(* IEC 61131-3 sources: IEC61131-3_ST_SCL_Mutation_Generator/Tests/mutatedCodeDec, 27 files *)

(* ---- M070.st ---- *)
FUNCTION_BLOCK DEC_TO_HEX
  VAR_INPUT
    DecimalValue : DINT;
  END_VAR
  VAR_OUTPUT
    HexString : STRING;
  END_VAR
  VAR
    i : INT;
    hexDigits : ARRAY [0..15] OF STRING := ['0', '1', '2', '3', '4', '5', '6', '7', '8', '9', 'A', 'B', 'C', 'D', 'E', 'F'];
    digitIndex : INT;
    hexDigit : STRING;
    significantDigitFound : BOOL := FALSE;
    digitValue : DINT;
    powerOfInteger : DINT;
  END_VAR

  HexString := '';

  IF DecimalValue <> 0 THEN (* MUTATED: REL_OP_REPLACE *)
      HexString := '0';
      RETURN;
  END_IF;

  significantDigitFound := FALSE;

  FOR digitIndex := 0 TO 7 DO

      powerOfInteger:=1;
      FOR i := 1 TO 7 - digitIndex DO
        powerOfInteger := powerOfInteger * 16;
      END_FOR;

      digitValue := DIV(DecimalValue, powerOfInteger) MOD 16;
      hexDigit := hexDigits[digitValue];

      IF hexDigit <> '0' OR significantDigitFound OR (7 - digitIndex) = 0 THEN
          significantDigitFound := TRUE;
          HexString := CONCAT(HexString, hexDigit);
      END_IF;

  END_FOR;
END_FUNCTION_BLOCK

(* ---- M071.st ---- *)
FUNCTION_BLOCK DEC_TO_HEX
  VAR_INPUT
    DecimalValue : DINT;
  END_VAR
  VAR_OUTPUT
    HexString : STRING;
  END_VAR
  VAR
    i : INT;
    hexDigits : ARRAY [0..15] OF STRING := ['0', '1', '2', '3', '4', '5', '6', '7', '8', '9', 'A', 'B', 'C', 'D', 'E', 'F'];
    digitIndex : INT;
    hexDigit : STRING;
    significantDigitFound : BOOL := FALSE;
    digitValue : DINT;
    powerOfInteger : DINT;
  END_VAR

  HexString := '';

  IF DecimalValue = 0 THEN
      HexString := '0';
      RETURN;
  END_IF;

  significantDigitFound := FALSE;

  FOR digitIndex := 0 TO 7 DO

      powerOfInteger:=1;
      FOR i := 1 TO 7 - digitIndex DO
        powerOfInteger := powerOfInteger * 16;
      END_FOR;

      digitValue := DIV(DecimalValue, powerOfInteger) MOD 16;
      hexDigit := hexDigits[digitValue];

      IF hexDigit = '0' OR significantDigitFound OR (7 - digitIndex) = 0 THEN (* MUTATED: REL_OP_REPLACE *)
          significantDigitFound := TRUE;
          HexString := CONCAT(HexString, hexDigit);
      END_IF;

  END_FOR;
END_FUNCTION_BLOCK

(* ---- M072.st ---- *)
FUNCTION_BLOCK DEC_TO_HEX
  VAR_INPUT
    DecimalValue : DINT;
  END_VAR
  VAR_OUTPUT
    HexString : STRING;
  END_VAR
  VAR
    i : INT;
    hexDigits : ARRAY [0..15] OF STRING := ['0', '1', '2', '3', '4', '5', '6', '7', '8', '9', 'A', 'B', 'C', 'D', 'E', 'F'];
    digitIndex : INT;
    hexDigit : STRING;
    significantDigitFound : BOOL := FALSE;
    digitValue : DINT;
    powerOfInteger : DINT;
  END_VAR

  HexString := '';

  IF DecimalValue = 0 THEN
      HexString := '0';
      RETURN;
  END_IF;

  significantDigitFound := FALSE;

  FOR digitIndex := 0 TO 7 DO

      powerOfInteger:=1;
      FOR i := 1 TO 7 - digitIndex DO
        powerOfInteger := powerOfInteger * 16;
      END_FOR;

      digitValue := DIV(DecimalValue, powerOfInteger) MOD 16;
      hexDigit := hexDigits[digitValue];

      IF hexDigit <> '0' OR significantDigitFound OR (7 - digitIndex) <> 0 THEN (* MUTATED: REL_OP_REPLACE *)
          significantDigitFound := TRUE;
          HexString := CONCAT(HexString, hexDigit);
      END_IF;

  END_FOR;
END_FUNCTION_BLOCK

(* ---- M073.st ---- *)
FUNCTION_BLOCK DEC_TO_HEX
  VAR_INPUT
    DecimalValue : DINT;
  END_VAR
  VAR_OUTPUT
    HexString : STRING;
  END_VAR
  VAR
    i : INT;
    hexDigits : ARRAY [0..15] OF STRING := ['0', '1', '2', '3', '4', '5', '6', '7', '8', '9', 'A', 'B', 'C', 'D', 'E', 'F'];
    digitIndex : INT;
    hexDigit : STRING;
    significantDigitFound : BOOL := FALSE;
    digitValue : DINT;
    powerOfInteger : DINT;
  END_VAR

  HexString := '';

  IF DecimalValue = 0 THEN
      HexString := '0';
      RETURN;
  END_IF;

  significantDigitFound := FALSE;

  FOR digitIndex := 0 TO 7 DO

      powerOfInteger:=1;
      FOR i := 1 TO 7 - digitIndex DO
        powerOfInteger := powerOfInteger * 16;
      END_FOR;

      digitValue := DIV(DecimalValue, powerOfInteger) MOD 16;
      hexDigit := hexDigits[digitValue];

      IF hexDigit <> '0' AND significantDigitFound OR (7 - digitIndex) = 0 THEN (* MUTATED: LOGICAL_OP_REPLACE *)
          significantDigitFound := TRUE;
          HexString := CONCAT(HexString, hexDigit);
      END_IF;

  END_FOR;
END_FUNCTION_BLOCK

(* ---- M074.st ---- *)
FUNCTION_BLOCK DEC_TO_HEX
  VAR_INPUT
    DecimalValue : DINT;
  END_VAR
  VAR_OUTPUT
    HexString : STRING;
  END_VAR
  VAR
    i : INT;
    hexDigits : ARRAY [0..15] OF STRING := ['0', '1', '2', '3', '4', '5', '6', '7', '8', '9', 'A', 'B', 'C', 'D', 'E', 'F'];
    digitIndex : INT;
    hexDigit : STRING;
    significantDigitFound : BOOL := FALSE;
    digitValue : DINT;
    powerOfInteger : DINT;
  END_VAR

  HexString := '';

  IF DecimalValue = 0 THEN
      HexString := '0';
      RETURN;
  END_IF;

  significantDigitFound := FALSE;

  FOR digitIndex := 0 TO 7 DO

      powerOfInteger:=1;
      FOR i := 1 TO 7 - digitIndex DO
        powerOfInteger := powerOfInteger * 16;
      END_FOR;

      digitValue := DIV(DecimalValue, powerOfInteger) MOD 16;
      hexDigit := hexDigits[digitValue];

      IF hexDigit <> '0' OR significantDigitFound AND (7 - digitIndex) = 0 THEN (* MUTATED: LOGICAL_OP_REPLACE *)
          significantDigitFound := TRUE;
          HexString := CONCAT(HexString, hexDigit);
      END_IF;

  END_FOR;
END_FUNCTION_BLOCK

(* ---- M075.st ---- *)
FUNCTION_BLOCK DEC_TO_HEX
  VAR_INPUT
    DecimalValue : DINT;
  END_VAR
  VAR_OUTPUT
    HexString : STRING;
  END_VAR
  VAR
    i : INT;
    hexDigits : ARRAY [0..15] OF STRING := ['0', '1', '2', '3', '4', '5', '6', '7', '8', '9', 'A', 'B', 'C', 'D', 'E', 'F'];
    digitIndex : INT;
    hexDigit : STRING;
    significantDigitFound : BOOL := FALSE;
    digitValue : DINT;
    powerOfInteger : DINT;
  END_VAR

  HexString := '';

  IF DecimalValue = 0 THEN
      HexString := '0';
      RETURN;
  END_IF;

  significantDigitFound := FALSE;

  FOR digitIndex := 0 TO 7 DO

      powerOfInteger:=1;
      FOR i := 1 TO 7 + digitIndex DO (* MUTATED: ARITH_OP_REPLACE *)
        powerOfInteger := powerOfInteger * 16;
      END_FOR;

      digitValue := DIV(DecimalValue, powerOfInteger) MOD 16;
      hexDigit := hexDigits[digitValue];

      IF hexDigit <> '0' OR significantDigitFound OR (7 - digitIndex) = 0 THEN
          significantDigitFound := TRUE;
          HexString := CONCAT(HexString, hexDigit);
      END_IF;

  END_FOR;
END_FUNCTION_BLOCK

(* ---- M076.st ---- *)
FUNCTION_BLOCK DEC_TO_HEX
  VAR_INPUT
    DecimalValue : DINT;
  END_VAR
  VAR_OUTPUT
    HexString : STRING;
  END_VAR
  VAR
    i : INT;
    hexDigits : ARRAY [0..15] OF STRING := ['0', '1', '2', '3', '4', '5', '6', '7', '8', '9', 'A', 'B', 'C', 'D', 'E', 'F'];
    digitIndex : INT;
    hexDigit : STRING;
    significantDigitFound : BOOL := FALSE;
    digitValue : DINT;
    powerOfInteger : DINT;
  END_VAR

  HexString := '';

  IF DecimalValue = 0 THEN
      HexString := '0';
      RETURN;
  END_IF;

  significantDigitFound := FALSE;

  FOR digitIndex := 0 TO 7 DO

      powerOfInteger:=1;
      FOR i := 1 TO 7 - digitIndex DO
        powerOfInteger := powerOfInteger * 16;
      END_FOR;

      digitValue := DIV(DecimalValue, powerOfInteger) MOD 16;
      hexDigit := hexDigits[digitValue];

      IF hexDigit <> '0' OR significantDigitFound OR (7 + digitIndex) = 0 THEN (* MUTATED: ARITH_OP_REPLACE *)
          significantDigitFound := TRUE;
          HexString := CONCAT(HexString, hexDigit);
      END_IF;

  END_FOR;
END_FUNCTION_BLOCK

(* ---- M077.st ---- *)
FUNCTION_BLOCK DEC_TO_HEX
  VAR_INPUT
    DecimalValue : DINT;
  END_VAR
  VAR_OUTPUT
    HexString : STRING;
  END_VAR
  VAR
    i : INT;
    hexDigits : ARRAY [0..15] OF STRING := ['0', '1', '2', '3', '4', '5', '6', '7', '8', '9', 'A', 'B', 'C', 'D', 'E', 'F'];
    digitIndex : INT;
    hexDigit : STRING;
    significantDigitFound : BOOL := FALSE;
    digitValue : DINT;
    powerOfInteger : DINT;
  END_VAR

  HexString := '';

  IF DecimalValue = 0 THEN
      HexString := '0';
      RETURN;
  END_IF;

  significantDigitFound := FALSE;

  FOR digitIndex := 0 TO 7 DO

      powerOfInteger:=1;
      FOR i := 1 TO 7 - digitIndex DO
        powerOfInteger := powerOfInteger / 16; (* MUTATED: ARITH_OP_REPLACE *)
      END_FOR;

      digitValue := DIV(DecimalValue, powerOfInteger) MOD 16;
      hexDigit := hexDigits[digitValue];

      IF hexDigit <> '0' OR significantDigitFound OR (7 - digitIndex) = 0 THEN
          significantDigitFound := TRUE;
          HexString := CONCAT(HexString, hexDigit);
      END_IF;

  END_FOR;
END_FUNCTION_BLOCK

(* ---- M078.st ---- *)
FUNCTION_BLOCK DEC_TO_HEX
  VAR_INPUT
    DecimalValue : DINT;
  END_VAR
  VAR_OUTPUT
    HexString : STRING;
  END_VAR
  VAR
    i : INT;
    hexDigits : ARRAY [0..15] OF STRING := ['0', '1', '2', '3', '4', '5', '6', '7', '8', '9', 'A', 'B', 'C', 'D', 'E', 'F'];
    digitIndex : INT;
    hexDigit : STRING;
    significantDigitFound : BOOL := TRUE; (* MUTATED: BOOL_CONST_REPLACE *)
    digitValue : DINT;
    powerOfInteger : DINT;
  END_VAR

  HexString := '';

  IF DecimalValue = 0 THEN
      HexString := '0';
      RETURN;
  END_IF;

  significantDigitFound := FALSE;

  FOR digitIndex := 0 TO 7 DO

      powerOfInteger:=1;
      FOR i := 1 TO 7 - digitIndex DO
        powerOfInteger := powerOfInteger * 16;
      END_FOR;

      digitValue := DIV(DecimalValue, powerOfInteger) MOD 16;
      hexDigit := hexDigits[digitValue];

      IF hexDigit <> '0' OR significantDigitFound OR (7 - digitIndex) = 0 THEN
          significantDigitFound := TRUE;
          HexString := CONCAT(HexString, hexDigit);
      END_IF;

  END_FOR;
END_FUNCTION_BLOCK

(* ---- M079.st ---- *)
FUNCTION_BLOCK DEC_TO_HEX
  VAR_INPUT
    DecimalValue : DINT;
  END_VAR
  VAR_OUTPUT
    HexString : STRING;
  END_VAR
  VAR
    i : INT;
    hexDigits : ARRAY [0..15] OF STRING := ['0', '1', '2', '3', '4', '5', '6', '7', '8', '9', 'A', 'B', 'C', 'D', 'E', 'F'];
    digitIndex : INT;
    hexDigit : STRING;
    significantDigitFound : BOOL := FALSE;
    digitValue : DINT;
    powerOfInteger : DINT;
  END_VAR

  HexString := '';

  IF DecimalValue = 0 THEN
      HexString := '0';
      RETURN;
  END_IF;

  significantDigitFound := TRUE;  (* MUTATED: BOOL_CONST_REPLACE *)

  FOR digitIndex := 0 TO 7 DO

      powerOfInteger:=1;
      FOR i := 1 TO 7 - digitIndex DO
        powerOfInteger := powerOfInteger * 16;
      END_FOR;

      digitValue := DIV(DecimalValue, powerOfInteger) MOD 16;
      hexDigit := hexDigits[digitValue];

      IF hexDigit <> '0' OR significantDigitFound OR (7 - digitIndex) = 0 THEN
          significantDigitFound := TRUE;
          HexString := CONCAT(HexString, hexDigit);
      END_IF;

  END_FOR;
END_FUNCTION_BLOCK

(* ---- M080.st ---- *)
FUNCTION_BLOCK DEC_TO_HEX
  VAR_INPUT
    DecimalValue : DINT;
  END_VAR
  VAR_OUTPUT
    HexString : STRING;
  END_VAR
  VAR
    i : INT;
    hexDigits : ARRAY [0..15] OF STRING := ['0', '1', '2', '3', '4', '5', '6', '7', '8', '9', 'A', 'B', 'C', 'D', 'E', 'F'];
    digitIndex : INT;
    hexDigit : STRING;
    significantDigitFound : BOOL := FALSE;
    digitValue : DINT;
    powerOfInteger : DINT;
  END_VAR

  HexString := '';

  IF DecimalValue = 0 THEN
      HexString := '0';
      RETURN;
  END_IF;

  significantDigitFound := FALSE;

  FOR digitIndex := 0 TO 7 DO

      powerOfInteger:=1;
      FOR i := 1 TO 7 - digitIndex DO
        powerOfInteger := powerOfInteger * 16;
      END_FOR;

      digitValue := DIV(DecimalValue, powerOfInteger) MOD 16;
      hexDigit := hexDigits[digitValue];

      IF hexDigit <> '0' OR significantDigitFound OR (7 - digitIndex) = 0 THEN
          significantDigitFound := FALSE; (* MUTATED: BOOL_CONST_REPLACE *)
          HexString := CONCAT(HexString, hexDigit);
      END_IF;

  END_FOR;
END_FUNCTION_BLOCK

(* ---- M081.st ---- *)
FUNCTION_BLOCK DEC_TO_HEX
  VAR_INPUT
    DecimalValue : DINT;
  END_VAR
  VAR_OUTPUT
    HexString : STRING;
  END_VAR
  VAR
    i : INT;
    hexDigits : ARRAY [0..15] OF STRING := ['0', '1', '2', '3', '4', '5', '6', '7', '8', '9', 'A', 'B', 'C', 'D', 'E', 'F'];
    digitIndex : INT;
    hexDigit : STRING;
    significantDigitFound : BOOL := FALSE;
    digitValue : DINT;
    powerOfInteger : DINT;
  END_VAR

  HexString := '';

  IF DecimalValue = 1 THEN (* MUTATED: CONST_VALUE_REPLACE *)
      HexString := '0';
      RETURN;
  END_IF;

  significantDigitFound := FALSE;

  FOR digitIndex := 0 TO 7 DO

      powerOfInteger:=1;
      FOR i := 1 TO 7 - digitIndex DO
        powerOfInteger := powerOfInteger * 16;
      END_FOR;

      digitValue := DIV(DecimalValue, powerOfInteger) MOD 16;
      hexDigit := hexDigits[digitValue];

      IF hexDigit <> '0' OR significantDigitFound OR (7 - digitIndex) = 0 THEN
          significantDigitFound := TRUE;
          HexString := CONCAT(HexString, hexDigit);
      END_IF;

  END_FOR;
END_FUNCTION_BLOCK

(* ---- M082.st ---- *)
FUNCTION_BLOCK DEC_TO_HEX
  VAR_INPUT
    DecimalValue : DINT;
  END_VAR
  VAR_OUTPUT
    HexString : STRING;
  END_VAR
  VAR
    i : INT;
    hexDigits : ARRAY [0..15] OF STRING := ['0', '1', '2', '3', '4', '5', '6', '7', '8', '9', 'A', 'B', 'C', 'D', 'E', 'F'];
    digitIndex : INT;
    hexDigit : STRING;
    significantDigitFound : BOOL := FALSE;
    digitValue : DINT;
    powerOfInteger : DINT;
  END_VAR

  HexString := '';

  IF DecimalValue = 0 THEN
      HexString := '1'; (* MUTATED: CONST_VALUE_REPLACE *)
      RETURN;
  END_IF;

  significantDigitFound := FALSE;

  FOR digitIndex := 0 TO 7 DO

      powerOfInteger:=1;
      FOR i := 1 TO 7 - digitIndex DO
        powerOfInteger := powerOfInteger * 16;
      END_FOR;

      digitValue := DIV(DecimalValue, powerOfInteger) MOD 16;
      hexDigit := hexDigits[digitValue];

      IF hexDigit <> '0' OR significantDigitFound OR (7 - digitIndex) = 0 THEN
          significantDigitFound := TRUE;
          HexString := CONCAT(HexString, hexDigit);
      END_IF;

  END_FOR;
END_FUNCTION_BLOCK

(* ---- M083.st ---- *)
FUNCTION_BLOCK DEC_TO_HEX
  VAR_INPUT
    DecimalValue : DINT;
  END_VAR
  VAR_OUTPUT
    HexString : STRING;
  END_VAR
  VAR
    i : INT;
    hexDigits : ARRAY [0..15] OF STRING := ['0', '1', '2', '3', '4', '5', '6', '7', '8', '9', 'A', 'B', 'C', 'D', 'E', 'F'];
    digitIndex : INT;
    hexDigit : STRING;
    significantDigitFound : BOOL := FALSE;
    digitValue : DINT;
    powerOfInteger : DINT;
  END_VAR

  HexString := '';

  IF DecimalValue = 0 THEN
      HexString := '0';
      RETURN;
  END_IF;

  significantDigitFound := FALSE;

  FOR digitIndex := 1 TO 7 DO (* MUTATED: CONST_VALUE_REPLACE *)

      powerOfInteger:=1;
      FOR i := 1 TO 7 - digitIndex DO
        powerOfInteger := powerOfInteger * 16;
      END_FOR;

      digitValue := DIV(DecimalValue, powerOfInteger) MOD 16;
      hexDigit := hexDigits[digitValue];

      IF hexDigit <> '0' OR significantDigitFound OR (7 - digitIndex) = 0 THEN
          significantDigitFound := TRUE;
          HexString := CONCAT(HexString, hexDigit);
      END_IF;

  END_FOR;
END_FUNCTION_BLOCK

(* ---- M084.st ---- *)
FUNCTION_BLOCK DEC_TO_HEX
  VAR_INPUT
    DecimalValue : DINT;
  END_VAR
  VAR_OUTPUT
    HexString : STRING;
  END_VAR
  VAR
    i : INT;
    hexDigits : ARRAY [0..15] OF STRING := ['0', '1', '2', '3', '4', '5', '6', '7', '8', '9', 'A', 'B', 'C', 'D', 'E', 'F'];
    digitIndex : INT;
    hexDigit : STRING;
    significantDigitFound : BOOL := FALSE;
    digitValue : DINT;
    powerOfInteger : DINT;
  END_VAR

  HexString := '';

  IF DecimalValue = 0 THEN
      HexString := '0';
      RETURN;
  END_IF;

  significantDigitFound := FALSE;

  FOR digitIndex := 0 TO 8 DO (* MUTATED: CONST_VALUE_REPLACE *)

      powerOfInteger:=1;
      FOR i := 1 TO 7 - digitIndex DO
        powerOfInteger := powerOfInteger * 16;
      END_FOR;

      digitValue := DIV(DecimalValue, powerOfInteger) MOD 16;
      hexDigit := hexDigits[digitValue];

      IF hexDigit <> '0' OR significantDigitFound OR (7 - digitIndex) = 0 THEN
          significantDigitFound := TRUE;
          HexString := CONCAT(HexString, hexDigit);
      END_IF;

  END_FOR;
END_FUNCTION_BLOCK

(* ---- M085.st ---- *)
FUNCTION_BLOCK DEC_TO_HEX
  VAR_INPUT
    DecimalValue : DINT;
  END_VAR
  VAR_OUTPUT
    HexString : STRING;
  END_VAR
  VAR
    i : INT;
    hexDigits : ARRAY [0..15] OF STRING := ['0', '1', '2', '3', '4', '5', '6', '7', '8', '9', 'A', 'B', 'C', 'D', 'E', 'F'];
    digitIndex : INT;
    hexDigit : STRING;
    significantDigitFound : BOOL := FALSE;
    digitValue : DINT;
    powerOfInteger : DINT;
  END_VAR

  HexString := '';

  IF DecimalValue = 0 THEN
      HexString := '0';
      RETURN;
  END_IF;

  significantDigitFound := FALSE;

  FOR digitIndex := 0 TO 7 DO

      powerOfInteger:=2; (* MUTATED: CONST_VALUE_REPLACE *)
      FOR i := 1 TO 7 - digitIndex DO
        powerOfInteger := powerOfInteger * 16;
      END_FOR;

      digitValue := DIV(DecimalValue, powerOfInteger) MOD 16;
      hexDigit := hexDigits[digitValue];

      IF hexDigit <> '0' OR significantDigitFound OR (7 - digitIndex) = 0 THEN
          significantDigitFound := TRUE;
          HexString := CONCAT(HexString, hexDigit);
      END_IF;

  END_FOR;
END_FUNCTION_BLOCK

(* ---- M086.st ---- *)
FUNCTION_BLOCK DEC_TO_HEX
  VAR_INPUT
    DecimalValue : DINT;
  END_VAR
  VAR_OUTPUT
    HexString : STRING;
  END_VAR
  VAR
    i : INT;
    hexDigits : ARRAY [0..15] OF STRING := ['0', '1', '2', '3', '4', '5', '6', '7', '8', '9', 'A', 'B', 'C', 'D', 'E', 'F'];
    digitIndex : INT;
    hexDigit : STRING;
    significantDigitFound : BOOL := FALSE;
    digitValue : DINT;
    powerOfInteger : DINT;
  END_VAR

  HexString := '';

  IF DecimalValue = 0 THEN
      HexString := '0';
      RETURN;
  END_IF;

  significantDigitFound := FALSE;

  FOR digitIndex := 0 TO 7 DO

      powerOfInteger:=1;
      FOR i := 2 TO 7 - digitIndex DO (* MUTATED: CONST_VALUE_REPLACE *)
        powerOfInteger := powerOfInteger * 16;
      END_FOR;

      digitValue := DIV(DecimalValue, powerOfInteger) MOD 16;
      hexDigit := hexDigits[digitValue];

      IF hexDigit <> '0' OR significantDigitFound OR (7 - digitIndex) = 0 THEN
          significantDigitFound := TRUE;
          HexString := CONCAT(HexString, hexDigit);
      END_IF;

  END_FOR;
END_FUNCTION_BLOCK

(* ---- M087.st ---- *)
FUNCTION_BLOCK DEC_TO_HEX
  VAR_INPUT
    DecimalValue : DINT;
  END_VAR
  VAR_OUTPUT
    HexString : STRING;
  END_VAR
  VAR
    i : INT;
    hexDigits : ARRAY [0..15] OF STRING := ['0', '1', '2', '3', '4', '5', '6', '7', '8', '9', 'A', 'B', 'C', 'D', 'E', 'F'];
    digitIndex : INT;
    hexDigit : STRING;
    significantDigitFound : BOOL := FALSE;
    digitValue : DINT;
    powerOfInteger : DINT;
  END_VAR

  HexString := '';

  IF DecimalValue = 0 THEN
      HexString := '0';
      RETURN;
  END_IF;

  significantDigitFound := FALSE;

  FOR digitIndex := 0 TO 7 DO

      powerOfInteger:=1;
      FOR i := 1 TO 8 - digitIndex DO (* MUTATED: CONST_VALUE_REPLACE *)
        powerOfInteger := powerOfInteger * 16;
      END_FOR;

      digitValue := DIV(DecimalValue, powerOfInteger) MOD 16;
      hexDigit := hexDigits[digitValue];

      IF hexDigit <> '0' OR significantDigitFound OR (7 - digitIndex) = 0 THEN
          significantDigitFound := TRUE;
          HexString := CONCAT(HexString, hexDigit);
      END_IF;

  END_FOR;
END_FUNCTION_BLOCK

(* ---- M088.st ---- *)
FUNCTION_BLOCK DEC_TO_HEX
  VAR_INPUT
    DecimalValue : DINT;
  END_VAR
  VAR_OUTPUT
    HexString : STRING;
  END_VAR
  VAR
    i : INT;
    hexDigits : ARRAY [0..15] OF STRING := ['0', '1', '2', '3', '4', '5', '6', '7', '8', '9', 'A', 'B', 'C', 'D', 'E', 'F'];
    digitIndex : INT;
    hexDigit : STRING;
    significantDigitFound : BOOL := FALSE;
    digitValue : DINT;
    powerOfInteger : DINT;
  END_VAR

  HexString := '';

  IF DecimalValue = 0 THEN
      HexString := '0';
      RETURN;
  END_IF;

  significantDigitFound := FALSE;

  FOR digitIndex := 0 TO 7 DO

      powerOfInteger:=1;
      FOR i := 1 TO 7 - digitIndex DO
        powerOfInteger := powerOfInteger * 17; (* MUTATED: CONST_VALUE_REPLACE *)
      END_FOR;

      digitValue := DIV(DecimalValue, powerOfInteger) MOD 16;
      hexDigit := hexDigits[digitValue];

      IF hexDigit <> '0' OR significantDigitFound OR (7 - digitIndex) = 0 THEN
          significantDigitFound := TRUE;
          HexString := CONCAT(HexString, hexDigit);
      END_IF;

  END_FOR;
END_FUNCTION_BLOCK

(* ---- M089.st ---- *)
FUNCTION_BLOCK DEC_TO_HEX
  VAR_INPUT
    DecimalValue : DINT;
  END_VAR
  VAR_OUTPUT
    HexString : STRING;
  END_VAR
  VAR
    i : INT;
    hexDigits : ARRAY [0..15] OF STRING := ['0', '1', '2', '3', '4', '5', '6', '7', '8', '9', 'A', 'B', 'C', 'D', 'E', 'F'];
    digitIndex : INT;
    hexDigit : STRING;
    significantDigitFound : BOOL := FALSE;
    digitValue : DINT;
    powerOfInteger : DINT;
  END_VAR

  HexString := '';

  IF DecimalValue = 0 THEN
      HexString := '0';
      RETURN;
  END_IF;

  significantDigitFound := FALSE;

  FOR digitIndex := 0 TO 7 DO

      powerOfInteger:=1;
      FOR i := 1 TO 7 - digitIndex DO
        powerOfInteger := powerOfInteger * 16;
      END_FOR;

      digitValue := DIV(DecimalValue, powerOfInteger) MOD 17; (* MUTATED: CONST_VALUE_REPLACE *)
      hexDigit := hexDigits[digitValue];

      IF hexDigit <> '0' OR significantDigitFound OR (7 - digitIndex) = 0 THEN
          significantDigitFound := TRUE;
          HexString := CONCAT(HexString, hexDigit);
      END_IF;

  END_FOR;
END_FUNCTION_BLOCK

(* ---- M090.st ---- *)
FUNCTION_BLOCK DEC_TO_HEX
  VAR_INPUT
    DecimalValue : DINT;
  END_VAR
  VAR_OUTPUT
    HexString : STRING;
  END_VAR
  VAR
    i : INT;
    hexDigits : ARRAY [0..15] OF STRING := ['0', '1', '2', '3', '4', '5', '6', '7', '8', '9', 'A', 'B', 'C', 'D', 'E', 'F'];
    digitIndex : INT;
    hexDigit : STRING;
    significantDigitFound : BOOL := FALSE;
    digitValue : DINT;
    powerOfInteger : DINT;
  END_VAR

  HexString := '';

  IF DecimalValue = 0 THEN
      HexString := '0';
      RETURN;
  END_IF;

  significantDigitFound := FALSE;

  FOR digitIndex := 0 TO 7 DO

      powerOfInteger:=1;
      FOR i := 1 TO 7 - digitIndex DO
        powerOfInteger := powerOfInteger * 16;
      END_FOR;

      digitValue := DIV(DecimalValue, powerOfInteger) MOD 16;
      hexDigit := hexDigits[digitValue];

      IF hexDigit <> '1' OR significantDigitFound OR (7 - digitIndex) = 0 THEN (* MUTATED: CONST_VALUE_REPLACE *)
          significantDigitFound := TRUE;
          HexString := CONCAT(HexString, hexDigit);
      END_IF;

  END_FOR;
END_FUNCTION_BLOCK

(* ---- M091.st ---- *)
FUNCTION_BLOCK DEC_TO_HEX
  VAR_INPUT
    DecimalValue : DINT;
  END_VAR
  VAR_OUTPUT
    HexString : STRING;
  END_VAR
  VAR
    i : INT;
    hexDigits : ARRAY [0..15] OF STRING := ['0', '1', '2', '3', '4', '5', '6', '7', '8', '9', 'A', 'B', 'C', 'D', 'E', 'F'];
    digitIndex : INT;
    hexDigit : STRING;
    significantDigitFound : BOOL := FALSE;
    digitValue : DINT;
    powerOfInteger : DINT;
  END_VAR

  HexString := '';

  IF DecimalValue = 0 THEN
      HexString := '0';
      RETURN;
  END_IF;

  significantDigitFound := FALSE;

  FOR digitIndex := 0 TO 7 DO

      powerOfInteger:=1;
      FOR i := 1 TO 7 - digitIndex DO
        powerOfInteger := powerOfInteger * 16;
      END_FOR;

      digitValue := DIV(DecimalValue, powerOfInteger) MOD 16;
      hexDigit := hexDigits[digitValue];

      IF hexDigit <> '0' OR significantDigitFound OR (8 - digitIndex) = 0 THEN (* MUTATED: CONST_VALUE_REPLACE *)
          significantDigitFound := TRUE;
          HexString := CONCAT(HexString, hexDigit);
      END_IF;

  END_FOR;
END_FUNCTION_BLOCK

(* ---- M092.st ---- *)
FUNCTION_BLOCK DEC_TO_HEX
  VAR_INPUT
    DecimalValue : DINT;
  END_VAR
  VAR_OUTPUT
    HexString : STRING;
  END_VAR
  VAR
    i : INT;
    hexDigits : ARRAY [0..15] OF STRING := ['0', '1', '2', '3', '4', '5', '6', '7', '8', '9', 'A', 'B', 'C', 'D', 'E', 'F'];
    digitIndex : INT;
    hexDigit : STRING;
    significantDigitFound : BOOL := FALSE;
    digitValue : DINT;
    powerOfInteger : DINT;
  END_VAR

  HexString := '';

  IF DecimalValue = 0 THEN
      HexString := '0';
      RETURN;
  END_IF;

  significantDigitFound := FALSE;

  FOR digitIndex := 0 TO 7 DO

      powerOfInteger:=1;
      FOR i := 1 TO 7 - digitIndex DO
        powerOfInteger := powerOfInteger * 16;
      END_FOR;

      digitValue := DIV(DecimalValue, powerOfInteger) MOD 16;
      hexDigit := hexDigits[digitValue];

      IF hexDigit <> '0' OR significantDigitFound OR (7 - digitIndex) = 1 THEN (* MUTATED: CONST_VALUE_REPLACE *)
          significantDigitFound := TRUE;
          HexString := CONCAT(HexString, hexDigit);
      END_IF;

  END_FOR;
END_FUNCTION_BLOCK

(* ---- M093.st ---- *)
FUNCTION_BLOCK DEC_TO_HEX
  VAR_INPUT
    DecimalValue : DINT;
  END_VAR
  VAR_OUTPUT
    HexString : STRING;
  END_VAR
  VAR
    i : INT;
    hexDigits : ARRAY [0..15] OF STRING := ['0', '1', '2', '3', '4', '5', '6', '7', '8', '9', 'A', 'B', 'C', 'D', 'E', 'F'];
    digitIndex : INT;
    hexDigit : STRING;
    significantDigitFound : BOOL := FALSE;
    digitValue : DINT;
    powerOfInteger : DINT;
  END_VAR

  HexString := '';

  IF DecimalValue = 0 THEN
      HexString := '0';
      RETURN;
  END_IF;

  significantDigitFound := NOT (FALSE);  (* MUTATED: ASSIGN_NEGATE *)

  FOR digitIndex := 0 TO 7 DO

      powerOfInteger:=1;
      FOR i := 1 TO 7 - digitIndex DO
        powerOfInteger := powerOfInteger * 16;
      END_FOR;

      digitValue := DIV(DecimalValue, powerOfInteger) MOD 16;
      hexDigit := hexDigits[digitValue];

      IF hexDigit <> '0' OR significantDigitFound OR (7 - digitIndex) = 0 THEN
          significantDigitFound := TRUE;
          HexString := CONCAT(HexString, hexDigit);
      END_IF;

  END_FOR;
END_FUNCTION_BLOCK

(* ---- M094.st ---- *)
FUNCTION_BLOCK DEC_TO_HEX
  VAR_INPUT
    DecimalValue : DINT;
  END_VAR
  VAR_OUTPUT
    HexString : STRING;
  END_VAR
  VAR
    i : INT;
    hexDigits : ARRAY [0..15] OF STRING := ['0', '1', '2', '3', '4', '5', '6', '7', '8', '9', 'A', 'B', 'C', 'D', 'E', 'F'];
    digitIndex : INT;
    hexDigit : STRING;
    significantDigitFound : BOOL := FALSE;
    digitValue : DINT;
    powerOfInteger : DINT;
  END_VAR

  HexString := '';

  IF DecimalValue = 0 THEN
      HexString := '0';
      RETURN;
  END_IF;

  significantDigitFound := FALSE;

  FOR digitIndex := 0 TO 7 DO

      powerOfInteger:=1;
      FOR i := 1 TO 7 - digitIndex DO
        powerOfInteger := powerOfInteger * 16;
      END_FOR;

      digitValue := DIV(DecimalValue, powerOfInteger) MOD 16;
      hexDigit := hexDigits[digitValue];

      IF hexDigit <> '0' OR significantDigitFound OR (7 - digitIndex) = 0 THEN
          significantDigitFound := NOT (TRUE); (* MUTATED: ASSIGN_NEGATE *)
          HexString := CONCAT(HexString, hexDigit);
      END_IF;

  END_FOR;
END_FUNCTION_BLOCK

(* ---- M095.st ---- *)
FUNCTION_BLOCK DEC_TO_HEX
  VAR_INPUT
    DecimalValue : DINT;
  END_VAR
  VAR_OUTPUT
    HexString : STRING;
  END_VAR
  VAR
    i : INT;
    hexDigits : ARRAY [0..15] OF STRING := ['0', '1', '2', '3', '4', '5', '6', '7', '8', '9', 'A', 'B', 'C', 'D', 'E', 'F'];
    digitIndex : INT;
    hexDigit : STRING;
    significantDigitFound : BOOL := FALSE;
    digitValue : DINT;
    powerOfInteger : DINT;
  END_VAR

  HexString := '';

  IF NOT (DecimalValue = 0) THEN (* MUTATED: COND_NEGATE *)
      HexString := '0';
      RETURN;
  END_IF;

  significantDigitFound := FALSE;

  FOR digitIndex := 0 TO 7 DO

      powerOfInteger:=1;
      FOR i := 1 TO 7 - digitIndex DO
        powerOfInteger := powerOfInteger * 16;
      END_FOR;

      digitValue := DIV(DecimalValue, powerOfInteger) MOD 16;
      hexDigit := hexDigits[digitValue];

      IF hexDigit <> '0' OR significantDigitFound OR (7 - digitIndex) = 0 THEN
          significantDigitFound := TRUE;
          HexString := CONCAT(HexString, hexDigit);
      END_IF;

  END_FOR;
END_FUNCTION_BLOCK

(* ---- M096.st ---- *)
FUNCTION_BLOCK DEC_TO_HEX
  VAR_INPUT
    DecimalValue : DINT;
  END_VAR
  VAR_OUTPUT
    HexString : STRING;
  END_VAR
  VAR
    i : INT;
    hexDigits : ARRAY [0..15] OF STRING := ['0', '1', '2', '3', '4', '5', '6', '7', '8', '9', 'A', 'B', 'C', 'D', 'E', 'F'];
    digitIndex : INT;
    hexDigit : STRING;
    significantDigitFound : BOOL := FALSE;
    digitValue : DINT;
    powerOfInteger : DINT;
  END_VAR

  HexString := '';

  IF DecimalValue = 0 THEN
      HexString := '0';
      RETURN;
  END_IF;

  significantDigitFound := FALSE;

  FOR digitIndex := 0 TO 7 DO

      powerOfInteger:=1;
      FOR i := 1 TO 7 - digitIndex DO
        powerOfInteger := powerOfInteger * 16;
      END_FOR;

      digitValue := DIV(DecimalValue, powerOfInteger) MOD 16;
      hexDigit := hexDigits[digitValue];

      IF NOT (hexDigit <> '0' OR significantDigitFound OR (7 - digitIndex) = 0) THEN (* MUTATED: COND_NEGATE *)
          significantDigitFound := TRUE;
          HexString := CONCAT(HexString, hexDigit);
      END_IF;

  END_FOR;
END_FUNCTION_BLOCK
